FUNCTION_BLOCK FTS_NCGenerator_Spy
VAR_IN_OUT
	stAxis: ST_Axis;
END_VAR
VAR_INPUT
	fCycleTime: LREAL;
END_VAR
VAR
	///_bCalStart             :BOOL:=FALSE;
	_bEnable: BOOL;
	///_bAutoPlan             :BOOL:=FALSE;
	_bCalculateDone: BOOL;
	_nIndex: UINT;
	_fLinearDealt: LREAL;
	_fLastPos: LREAL;
END_VAR
VAR CONSTANT
	cStateIdle: INT := 0;
	cStateReady: INT := 1;
	cStatePathGenerator: INT := 2;
	cDealtGap: REAL := 10000;
	cNcCycle: REAL := 0.001;
	cPointBuffer: UINT := 10;
END_VAR

// control logic 

IF stAxis.stPLCTONC.bNcEnable  THEN
 
   A_GetPosition();
ELSE
	stAxis.stAxisStatus.nNcCycleCounter:=0;
END_IF

ACTION A_GetPosition:


IF (stAxis.stPLCTONC.ePlanningMode=E_PlanningMode.PLANNINGMODE_LINEAR)THEN 
    A_LinearPosition();
ELSE
	;
END_IF
END_ACTION

ACTION A_LinearPosition:


stAxis.stAxisStatus.nNcCycleCounter:=stAxis.stAxisStatus.nNcCycleCounter+1;
IF (_fLastPos<>stAxis.stPLCTONC.stEndPosition.fPosition) THEN 
	IF (stAxis.stPLCTONC.nLinearPointNum<>0)THEN
        _fLinearDealt:=(stAxis.stPLCTONC.stEndPosition.fPosition-stAxis.stNcTOPLC.fActPos)/stAxis.stPLCTONC.nLinearPointNum;
	ELSE
		_fLinearDealt:=(stAxis.stPLCTONC.stEndPosition.fPosition-stAxis.stNcTOPLC.fActPos)/10;
	END_IF
END_IF 

	
stAxis.stNcTOPLC.fActPos:=stAxis.stNcTOPLC.fActPos+_fLinearDealt;	
stAxis.stNcTOPLC.fSetPos:=stAxis.stNcTOPLC.fActPos;


stAxis.stNcTOPLC.fSetVelo:=_fLinearDealt/0.001;
stAxis.stNcTOPLC.fActVelo:=_fLinearDealt/0.001;

IF (stAxis.stNcTOPLC.fActPos>=stAxis.stPLCTONC.stEndPosition.fPosition)THEN
	_fLinearDealt:=0;
END_IF

_fLastPos:=stAxis.stPLCTONC.stEndPosition.fPosition;
END_ACTION

END_FUNCTION_BLOCK

(* stored: Version 1.1.0.1, ProductVersion 3.1.4024.12
   POU FTS_NCGenerator_Spy: Id {54dc7b8d-25b6-4f55-8299-36f384b73c18}, SpecialFunc None
   Action A_GetPosition: Id {f8cefc2f-ba91-43a5-9460-08cd1e4551ea}
   Action A_LinearPosition: Id {c3a4d63f-417c-4e77-9b53-d54870472712} *)
